(* PLC project DeepSeek1.project, CODESYS CODESYS V3.5 SP20 *)
(* stored: creationDateTime 2026-10-15T18:39:41.03229, modificationDateTime 2026-10-15T18:34:13.9284842 *)

PROGRAM PLC_PRG
  VAR_INPUT
    i_bStart : BOOL;
    i_bStop : BOOL;
    i_wTempSensor : INT;
  END_VAR
  VAR_OUTPUT
    o_bHeater : BOOL;
    o_bMixer : BOOL;
    o_rAvgTemp : REAL;
  END_VAR
  VAR
    a_rTempHistory : ARRAY[1..5] OF REAL;
    fbMixTimer : TON;
    i_State : INT := 0;
    i_Index : INT;
    r_TempConverted : REAL;
    r_SumTemp : REAL;
    b_EmergencyStop : BOOL;
  END_VAR

                    
b_EmergencyStop := NOT i_bStop;

IF b_EmergencyStop THEN
    i_State := 0;
    fbMixTimer(IN := FALSE, PT := T#10S);
    o_bHeater := FALSE;
    o_bMixer := FALSE;
ELSE
    r_TempConverted := (INT_TO_REAL(i_wTempSensor) / 27648.0) * 150.0;

    FOR i_Index := 5 TO 2 BY -1 DO
        a_rTempHistory[i_Index] := a_rTempHistory[i_Index - 1];
    END_FOR;
    a_rTempHistory[1] := r_TempConverted;

    r_SumTemp := 0.0;
    FOR i_Index := 1 TO 5 DO
        r_SumTemp := r_SumTemp + a_rTempHistory[i_Index];
    END_FOR;
    o_rAvgTemp := r_SumTemp / 5.0;

    CASE i_State OF
        0:
            o_bHeater := FALSE;
            o_bMixer := FALSE;
            fbMixTimer(IN := FALSE, PT := T#10S);
            IF i_bStart THEN
                i_State := 1;
            END_IF;

        1:
            o_bHeater := TRUE;
            o_bMixer := FALSE;
            IF o_rAvgTemp > 80.0 THEN
                o_bHeater := FALSE;
                o_bMixer := TRUE;
                fbMixTimer(IN := TRUE, PT := T#10S);
                i_State := 2;
            END_IF;

        2:
            o_bHeater := FALSE;
            o_bMixer := TRUE;
            fbMixTimer(IN := TRUE, PT := T#10S);
            IF fbMixTimer.Q THEN
                o_bMixer := FALSE;
                fbMixTimer(IN := FALSE, PT := T#10S);
                i_State := 0;
            END_IF;

        ELSE
            i_State := 0;
            o_bHeater := FALSE;
            o_bMixer := FALSE;
    END_CASE;
END_IF;
                  
END_PROGRAM

CONFIGURATION Device
  RESOURCE Application ON PLC
    TASK MainTask(INTERVAL := T#20ms, PRIORITY := 1);
    PROGRAM PLC_PRG WITH MainTask : PLC_PRG;
  END_RESOURCE
END_CONFIGURATION
